(*
SPDX-FileCopyrightText: c 2026 Oleksandr Tiutyk <trofimich@gmail.com>
SPDX-License-Identifier: MIT
License: https://opensource.org/license/mit
*)

(*!
<summary>Checks scalar and short text formatting through the fitted ANY API.</summary>
<description>
Uses one task and stays at a stable address while assertions are bound to this instance.
</description>
*)

{attribute 'no_assign'}
{attribute 'no_explicit_call' := 'do not call this function block directly'}
FUNCTION_BLOCK WideStringFitFormattingTest EXTENDS TOF_Testing.SingleCycleTest
VAR_STAT
	{attribute 'hide'}
	_ClassName : STRING := __POUNAME();
END_VAR

(*!
<summary>Checks scalar and short text formatting through the fitted ANY API.</summary>
*)
METHOD PROTECTED ExecuteTest
VAR
	formatted : WSTRING(255);
	enabled : BOOL := TRUE;
	number : DINT := 12345;
	narrowText : STRING(50) := 'Sample string';
	wideText : WSTRING(50) := "Sample wide string";
END_VAR
formatted := TOF_Core.WideStrings.AnyToStringFit255(value := enabled);
Assert.ThatBool(
	actual := formatted = "TRUE",
	message := "AnyToStringFit255 must format BOOL"
).IsTrue();

formatted := TOF_Core.WideStrings.AnyToStringFit255(value := number);
Assert.ThatBool(
	actual := formatted = "12345",
	message := "AnyToStringFit255 must format DINT"
).IsTrue();

formatted := TOF_Core.WideStrings.AnyToStringFit255(value := narrowText);
Assert.ThatBool(
	actual := formatted = "Sample string",
	message := "AnyToStringFit255 must convert short STRING to WSTRING"
).IsTrue();

formatted := TOF_Core.WideStrings.AnyToStringFit255(value := wideText);
Assert.ThatBool(
	actual := formatted = "Sample wide string",
	message := "AnyToStringFit255 must pass short WSTRING as-is"
).IsTrue();
END_METHOD

//! <summary>Borrows the concrete class name. Callers must not modify it.</summary>
{attribute 'monitoring' := 'call'}
PROPERTY ClassName : REFERENCE TO STRING
GET
ClassName REF= _ClassName;
END_GET
END_PROPERTY

//! <summary>Borrows the compiler-initialized namespace name. Callers must not modify it.</summary>
{attribute 'monitoring' := 'call'}
PROPERTY NamespaceName : REFERENCE TO STRING
GET
NamespaceName REF= CurrentNamespace.Name;
END_GET
END_PROPERTY

//! <summary>Reports the concrete instance size in bytes.</summary>
{attribute 'monitoring' := 'call'}
PROPERTY SelfSize : ULINT
GET
SelfSize := XSIZEOF(THIS^);
END_GET
END_PROPERTY

END_FUNCTION_BLOCK

(* stored: Version 1.1.0.1
   POU WideStringFitFormattingTest: Id {fdce5f12-caf7-4f51-be4c-ccee78e39955}, SpecialFunc None
   Method ExecuteTest: Id {067c878a-361e-49db-a293-718cac03aacb}
   Property ClassName: Id {6849256d-822d-42f3-bbc8-eeb26e258427}
   Get Get: Id {57d0a892-8f65-4901-b684-387da06c2ada}
   Property NamespaceName: Id {ff95535c-6125-4f5c-afe1-e3ab627bfe62}
   Get Get: Id {44d3fd9f-f5d6-4ba7-8c20-6ac0ac4df9ea}
   Property SelfSize: Id {efd93286-4244-4528-a34a-83f5d657a132}
   Get Get: Id {6fb3af60-c3d2-474a-9a3c-5d78d04078f9} *)
